{attribute 'linkalways'}
{attribute 'no_explicit_call' := 'This FB is a CLASS and must be accessed using methods or properties'}
{attribute 'enable_dynamic_creation'}
FUNCTION_BLOCK Node_F_VN_InnerCircleExp EXTENDS VisionNode
VAR
    ipSrcImage : _ITcVnImage;
    fRadius : _LREAL(0.0);
    aCenter : _TcVnPoint2_REAL;
    eDistanceType : _ETcVnDistanceType(ETcVnDistanceType.TCVN_DT_L2);
    eMaskSize : _ETcVnDistanceTransformationMask(ETcVnDistanceTransformationMask.TCVN_DTM_5);
    hrPrev : _HRESULT(S_OK);
    hresult : _HRESULT(S_OK);
END_VAR

METHOD PUBLIC Clone : I_Node
VAR
    pNode : POINTER TO Node_F_VN_InnerCircleExp;
END_VAR
pNode := __NEW(Node_F_VN_InnerCircleExp);
Clone := pNode^;
END_METHOD

METHOD FB_init : BOOL
VAR_INPUT
    bInitRetains : BOOL;
    bInCopyCode : BOOL;
END_VAR
AddInput('ipSrcImage', ipSrcImage);
AddParameter('eDistanceType', eDistanceType);
AddParameter('eMaskSize', eMaskSize);
AddInput('hrPrev', hrPrev);
AddOutput('fRadius', fRadius);
AddOutput('aCenter', aCenter);
AddOutput('hresult', hresult);
END_METHOD

METHOD PROTECTED OnExecute
hresult.Value := F_VN_InnerCircleExp(
    ipSrcImage := ipSrcImage.Value,
    fRadius := fRadius.Value,
    aCenter := aCenter.Value,
    eDistanceType := eDistanceType.Value,
    eMaskSize := eMaskSize.Value,
    hrPrev := hrPrev.Value);
END_METHOD

METHOD PUBLIC PreExecutionCheck
VAR_INPUT
    Check : I_PreExecutionChecks;
END_VAR
VAR
    distanceTypeIsValid : BOOL;
END_VAR
Check.IsTrue(ipSrcImage.IsValid, 'ipSrcImage must contain an image');
Check.IsTrue(ipSrcImage.HasChannelCount(1), 'ipSrcImage must have 1 channel');
Check.IsTrue(ipSrcImage.IsElementType(ETcVnElementType.TCVN_ET_USINT), 'ipSrcImage must contain USINT elements');

CASE eDistanceType.Value OF
    ETcVnDistanceType.TCVN_DT_L1,
    ETcVnDistanceType.TCVN_DT_L2,
    ETcVnDistanceType.TCVN_DT_C :
        distanceTypeIsValid := TRUE;
END_CASE
Check.IsTrue(distanceTypeIsValid, 'eDistanceType value is unsupported');
END_METHOD

END_FUNCTION_BLOCK
